// TwinCAT 3 PLC project StudentPLC
// ProgramVersion: 3.1.4026.20
// libraries:
//   CmpBitmapPool, * (System)
//   Tc2_Standard, * (Beckhoff Automation GmbH)
//   Tc2_System, * (Beckhoff Automation GmbH)
//   Tc3_Module, * (Beckhoff Automation GmbH)
//   VisuSymbols,3.5.10.0,System
// project tree:
//   / GlobalTextList.TcGTLO, PlcTask.TcTTO, Visualization Manager.TcVMO (not stored)
//   GVLs/ GVLStudent.TcGVL
//   POUs/ LampDelay.TcPOU, LampStudent.TcPOU, LongHandshake.TcPOU, MAIN.TcPOU, RunStudent.TcPOU, ShortHandshake.TcPOU
//   VISUs/ VisualizationStudent.TcVIS
// real-time tasks:
//   TASK PlcTask: cycle T#10ms, priority 20, ADS port 350
//   TASK PlcTask1: cycle T#10ms, priority 21, ADS port 351
// variable links:
//   StudentPLC/StudentPLC Instance <-> slavePLC/slavePLC Instance
//     PlcTask Inputs/GVLStudent.ixStrobOne <-> PlcTask Outputs/GVLSlave.oxStrobOne
//     PlcTask Inputs/GVLStudent.ixStrobTwo <-> PlcTask Outputs/GVLSlave.oxStrobTwo
//     PlcTask Outputs/GVLStudent.IXButtonLong <-> PlcTask Inputs/GVLSlave.ixLong
//     PlcTask Outputs/GVLStudent.IXButtonShort <-> PlcTask Inputs/GVLSlave.ixShort
//     PlcTask Outputs/GVLStudent.oxStrobOne <-> PlcTask Inputs/GVLSlave.ixStrobOne
//     PlcTask Outputs/GVLStudent.oxStrobTwo <-> PlcTask Inputs/GVLSlave.ixStrobTwo

CONFIGURATION StudentPLC
    RESOURCE PLC ON TwinCAT3
        TASK PlcTask(INTERVAL := T#10ms, PRIORITY := 20);
        PROGRAM MAIN WITH PlcTask : MAIN;
    END_RESOURCE
END_CONFIGURATION

// ---- GVLs/GVLStudent.TcGVL
{attribute 'qualified_only'}
VAR_GLOBAL
	// Lamp varibols
	OXLampOXOne :BOOL;
	OXLampIXOneGreen :BOOL;
	OXLampOXTwo :BOOL;
	OXLampIXTwoGreen :BOOL;
	
	// Button varibols
	IXButtonShort AT %Q* :BOOL;
	IXButtonLong AT %Q*:BOOL;
	// strob out 
	oxStrobOne AT %Q* : BOOL ;
	oxStrobTwo AT %Q* : BOOL ;
 	// strob in
	ixStrobOne AT %I* : BOOL ;
	ixStrobTwo AT %I* : BOOL ; 
END_VAR

// ---- POUs/MAIN.TcPOU
PROGRAM MAIN
VAR
	
END_VAR

RunStudent();

END_PROGRAM

// ---- POUs/RunStudent.TcPOU
PROGRAM RunStudent
VAR
	LampStudent_0: LampStudent;
	ixStrobOne :BOOL;
	ixStrobTwo :BOOL;
	ixStrob: BOOL;
	LongHandshake_0: LongHandshake;
	ShortHandshake_0: ShortHandshake;
END_VAR

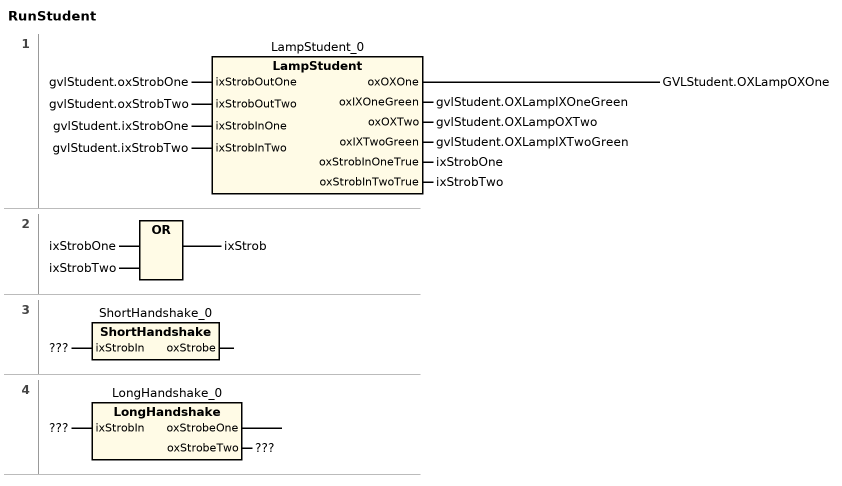
// NETWORK 1
LampStudent_0(
    ixStrobOutOne := gvlStudent.oxStrobOne,
    ixStrobOutTwo := gvlStudent.oxStrobTwo,
    ixStrobInOne := gvlStudent.ixStrobOne,
    ixStrobInTwo := gvlStudent.ixStrobTwo,
    oxIXOneGreen => gvlStudent.OXLampIXOneGreen,
    oxOXTwo => gvlStudent.OXLampOXTwo,
    oxIXTwoGreen => gvlStudent.OXLampIXTwoGreen,
    oxStrobInOneTrue => ixStrobOne,
    oxStrobInTwoTrue => ixStrobTwo); // LampStudent
GVLStudent.OXLampOXOne := LampStudent_0.oxOXOne;

// NETWORK 2
ixStrob := ixStrobOne OR ixStrobTwo;

// NETWORK 3
ShortHandshake_0(); // ShortHandshake

// NETWORK 4
LongHandshake_0(); // LongHandshake

END_PROGRAM

// ---- POUs/LampStudent.TcPOU
FUNCTION_BLOCK LampStudent
VAR_INPUT
	ixStrobOutOne :BOOL; // Direct control for group One main lamp (OX1)
	ixStrobOutTwo :BOOL; // Direct control for group Two main lamp (OX2)
	
	ixStrobInOne: BOOL; // Start signal for LampDelay sequence (group One)
	ixStrobInTwo: BOOL; // Start signal for LampDelay sequence (group Two)

END_VAR
VAR_OUTPUT
	  // Group One: main lamp + 3 indicator lamps (R, B, G)
	oxOXOne :BOOL; // Main lamp (direct)
	
	oxIXOneGreen :BOOL; // Indicator Green (from LampDelay)

	
	oxOXTwo :BOOL; // Main lamp (direct)
	
	oxIXTwoGreen :BOOL; // Indicator Green (from LampDelay)

	
	oxStrobInOneTrue: BOOL; // TRUE when all three indicators (group One) are ON
	oxStrobInTwoTrue: BOOL;// TRUE when all three indicators (group Two) are ON
	
END_VAR
	
VAR
	
	LampIXOne : LampDelay; // Instance for group One sequence
	LampIXTwo : LampDelay; // Instance for group Two sequence
	
END_VAR

// ------------------------------
// Direct main-lamp control
// ------------------------------

IF ixStrobOutOne THEN
	oxOXOne := TRUE;
ELSE
	oxOXOne := FALSE;
END_IF

IF ixStrobOutTwo THEN
	oxOXTwo := TRUE;
ELSE
	oxOXTwo := FALSE;
END_IF



// ------------------------------
// Group One: delayed indicator sequence
// ------------------------------
LampIXOne(ixStart := ixStrobInOne);

// Map LampDelay outputs to group One indicators

oxIXOneGreen     := LampIXOne.oxLampThree; // Green
oxStrobInOneTrue := LampIXOne.oxAllLightsOn; // All indicators ON


// ------------------------------
// Group Two: delayed indicator sequence
// ------------------------------
LampIXTwo(ixStart := ixStrobInTwo);

// Map LampDelay outputs to group Two indicators

oxIXTwoGreen     := LampIXTwo.oxLampThree; // Green
oxStrobInTwoTrue := LampIXTwo.oxAllLightsOn; // All indicators ON

END_FUNCTION_BLOCK

// ---- POUs/LampDelay.TcPOU
FUNCTION_BLOCK LampDelay
VAR_INPUT
    ixStart : BOOL;      // Start command: TRUE = run "power-up" sequence; FALSE = run "power-down" sequence
END_VAR
VAR_OUTPUT
    oxLampThree    : BOOL; // Output: Lamp 3 on/off
    oxAllLightsOn  : BOOL; // TRUE when all three lamps are on
END_VAR
VAR
    t      : TON;             // TON timer instance (non-retentive on IN falling edge)
    step   : INT := 0;        // State machine step
    delay  : TIME := T#150MS;    // Delay duration used between steps
    tStart : BOOL;            // Timer IN signal (acts like a "strobe" to start the TON)
    tEnd   : BOOL;            // TRUE when timer has elapsed (t.Q)
END_VAR


//_______________________________________________________________________________________________
// LampDelay is a step-sequenced (state machine) controller that turns on three lamps
// one BY one with a fixed delay between each stage when ixStart is TRUE. 
// When ixStart goes FALSE, it turns the lamps off again in reverse order, also with delays. 
// A TON timer (t) provides the per-step delay. oxAllLightsOn is TRUE once all three lamps are on.
//_______________________________________________________________________________________________


// ------------------------------
// State machine for sequenced on/off with delays
// ------------------------------
CASE step OF

    0: // Idle/reset: all lamps off, wait for start
        oxLampThree    := FALSE;
        oxAllLightsOn  := FALSE;
        IF ixStart THEN
            // Start power-up sequence: immediately turn on Lamp 1 and start delay
            tStart    := TRUE;                  // Start the TON for the next step delay
			t(IN := tStart, PT := delay);
            step      := 20;
        END_IF


    20: // After Lamp 2 is on, wait delay, then turn on Lamp 3
        IF tEnd THEN
            tStart := FALSE;                   // Reset TON input before next start
            t(IN := tStart, PT := delay);
            oxLampThree := TRUE;
            step := 30;
        END_IF

    30: // All three lamps are on; assert "all on" and wait for stop command
        oxAllLightsOn := TRUE;
        IF NOT ixStart THEN
            // Begin power-down sequence after stop command
            tStart := TRUE;                    // Start delay before turning lamps off
            t(IN := tStart, PT := delay);
            step := 60;
        END_IF


    60: // Wait delay, then turn off Lamp 1 and return to idle
        IF tEnd THEN
            oxLampThree := FALSE;
			tStart := FALSE;
			t(IN := tStart,  PT := delay);
            step := 0;                         // Back to idle
        END_IF

END_CASE

// ------------------------------
// Timer execution (must be called each cycle)
// ------------------------------
t(IN := tStart, PT := delay);  // Evaluate TON with current IN/PT
tEnd := t.Q;                   // Timer done flag for step logic

END_FUNCTION_BLOCK

// ---- POUs/LongHandshake.TcPOU
FUNCTION_BLOCK LongHandshake
VAR_INPUT
	ixStrobIn : BOOL;
END_VAR
VAR_OUTPUT
	oxStrobeOne : BOOL;
	oxStrobeTwo : BOOL;
END_VAR
VAR
END_VAR

END_FUNCTION_BLOCK

// ---- POUs/ShortHandshake.TcPOU
FUNCTION_BLOCK ShortHandshake
VAR_INPUT
	ixStrobIn : BOOL;
END_VAR
VAR_OUTPUT
	oxStrobe : BOOL;
END_VAR
VAR
END_VAR

END_FUNCTION_BLOCK

// ---- GlobalTextList.TcGTLO
TEXTLIST GlobalTextList
  378 = 'IXOne'
  913 = 'IXTwo'
  175 = 'loadding'
  693 = 'loading'
  725 = 'Long handshake'
  923 = 'Looding'
  572 = 'Master PLC'
  739 = 'Master strob one send'
  50 = 'Master strob two send'
  816 = 'OXOne'
  226 = 'OXTwo'
  198 = 'Short handshake'
  252 = 'Slav strob one send'
  968 = 'Strobe received'
  419 = 'This is student plc'
END_TEXTLIST

// ---- VISUs/VisualizationStudent.TcVIS
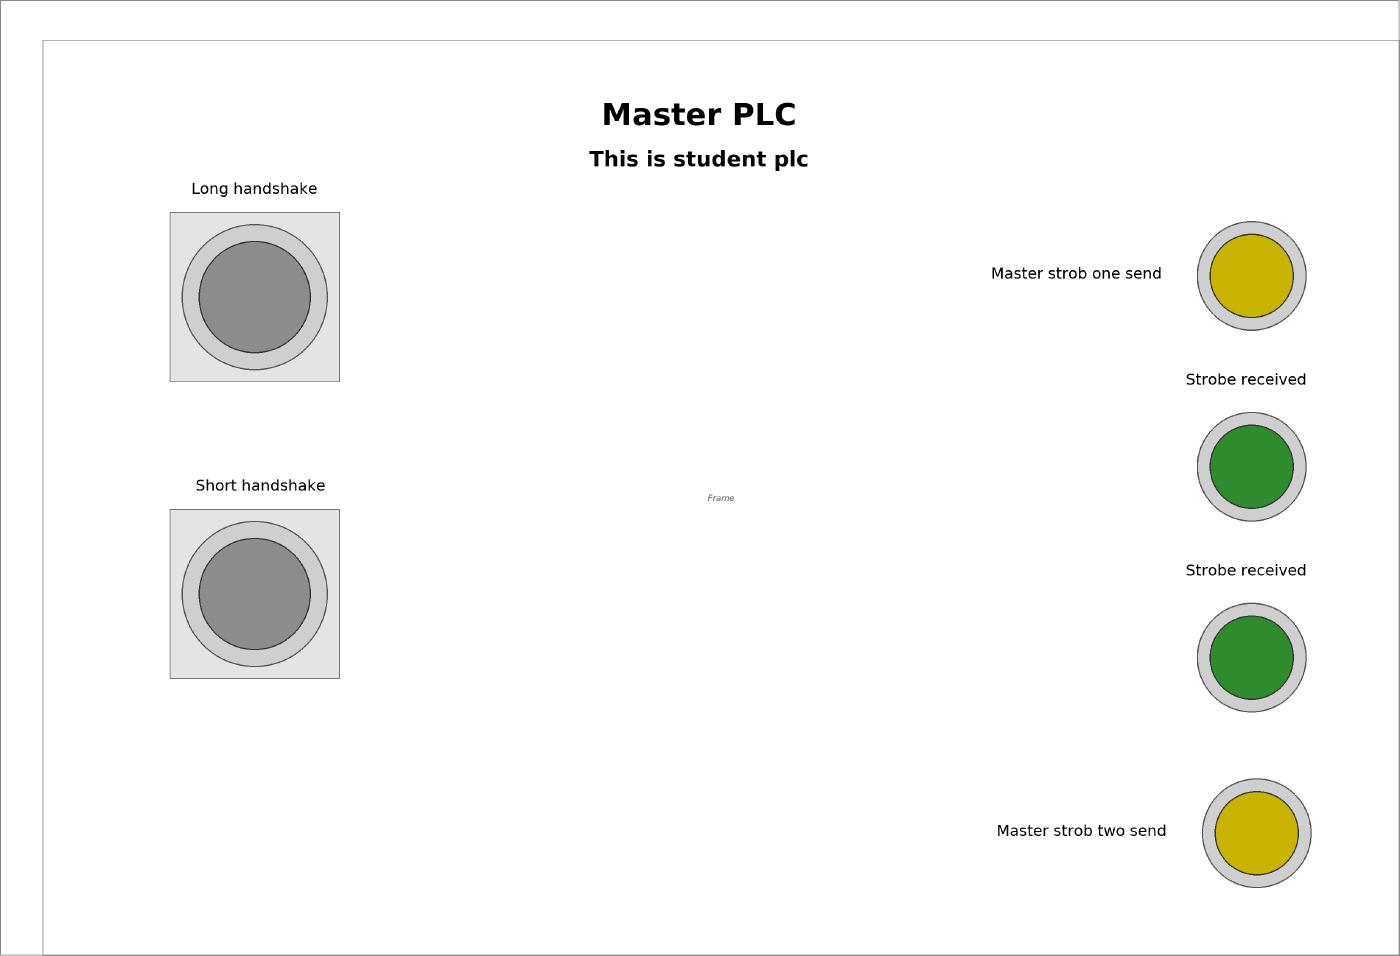
VISUALIZATION VisualizationStudent  // 1650x1127
    Frame (50,47 1600x1080)
    Label (699,110 250x50), "Master PLC"
    PushSwitch (200,250 200x200), variable: GVLStudent.IXButtonLong, behaviour: TAP, style: Switch-PushSwitch-Gray
    PushSwitch (200,600 200x200), variable: GVLStudent.IXButtonShort, behaviour: TAP, style: Switch-PushSwitch-Gray
    Label (225,200 150x45), "Long handshake"
    Label (225,550 164x45), "Short handshake"
    Label (1095,300 348x45), "Master strob one send"
    Lamp1 (1400,475 150x150), variable: GVLStudent.OXLampIXOneGreen, style: Lamp-Lamp1-Green
    Lamp1 (1406,907 150x150), variable: GVLStudent.OXLampOXTwo, style: Lamp-Lamp1-Yellow
    Lamp1 (1400,250 150x150), variable: GVLStudent.OXLampOXOne, style: Lamp-Lamp1-Yellow
    Label (1350,425 238x45), "Strobe received"
    Label (1101,957 348x45), "Master strob two send"
    Lamp1 (1400,700 150x150), variable: GVLStudent.OXLampIXTwoGreen, style: Lamp-Lamp1-Green
    Label (1350,650 238x45), "Strobe received"
    Label (643,172 362x30), "This is student plc"
END_VISUALIZATION
